Fanuc KAREL source: compact_preamble.KL

PROGRAM KB00003
%NOLOCKGROUP
VAR
P1:REAL;RESULT:REAL
BEGIN
P1=1.0
RESULT=ACOS(P1)
END KB00003
